// TIA Portal V20 export
ORGANIZATION_BLOCK "T7_Ciclo"   // OB130, LAD, ProgramCycle
TITLE = T7_Ciclo
{ S7_Optimized_Access := 'TRUE' }
AUTHOR : IA
FAMILY : PRUEBA
VERSION : 0.1
// Tanda 3: llama a todas las pruebas
// stored: AutoNumber false, IsIECCheckEnabled false, SetENOAutomatically false
   VAR_INPUT
      Initial_Call : Bool;
      Remanence : Bool;
   END_VAR
BEGIN

REGION Network 1: T7_Base
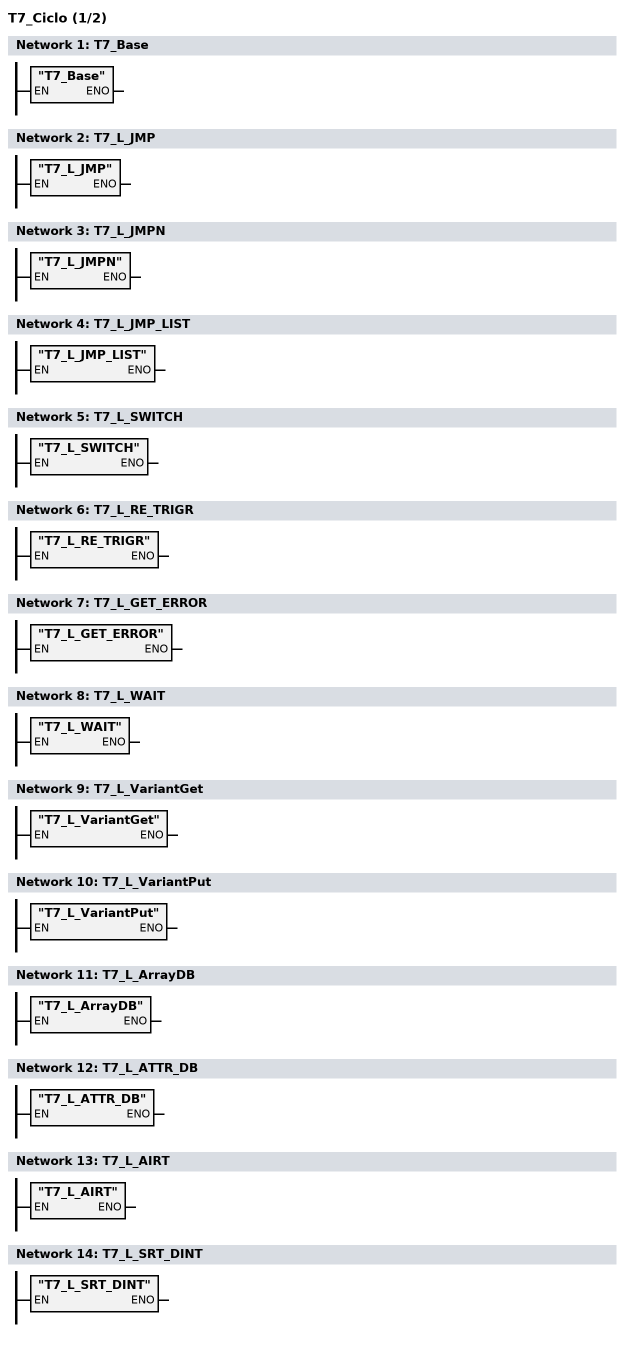
   RUNG wire#powerrail
      "T7_Base"()
   END_RUNG
   // the same network as SCL:
   "T7_Base"();
END_REGION

REGION Network 2: T7_L_JMP
   RUNG wire#powerrail
      "T7_L_JMP"()
   END_RUNG
   // the same network as SCL:
   "T7_L_JMP"();
END_REGION

REGION Network 3: T7_L_JMPN
   RUNG wire#powerrail
      "T7_L_JMPN"()
   END_RUNG
   // the same network as SCL:
   "T7_L_JMPN"();
END_REGION

REGION Network 4: T7_L_JMP_LIST
   RUNG wire#powerrail
      "T7_L_JMP_LIST"()
   END_RUNG
   // the same network as SCL:
   "T7_L_JMP_LIST"();
END_REGION

REGION Network 5: T7_L_SWITCH
   RUNG wire#powerrail
      "T7_L_SWITCH"()
   END_RUNG
   // the same network as SCL:
   "T7_L_SWITCH"();
END_REGION

REGION Network 6: T7_L_RE_TRIGR
   RUNG wire#powerrail
      "T7_L_RE_TRIGR"()
   END_RUNG
   // the same network as SCL:
   "T7_L_RE_TRIGR"();
END_REGION

REGION Network 7: T7_L_GET_ERROR
   RUNG wire#powerrail
      "T7_L_GET_ERROR"()
   END_RUNG
   // the same network as SCL:
   "T7_L_GET_ERROR"();
END_REGION

REGION Network 8: T7_L_WAIT
   RUNG wire#powerrail
      "T7_L_WAIT"()
   END_RUNG
   // the same network as SCL:
   "T7_L_WAIT"();
END_REGION

REGION Network 9: T7_L_VariantGet
   RUNG wire#powerrail
      "T7_L_VariantGet"()
   END_RUNG
   // the same network as SCL:
   "T7_L_VariantGet"();
END_REGION

REGION Network 10: T7_L_VariantPut
   RUNG wire#powerrail
      "T7_L_VariantPut"()
   END_RUNG
   // the same network as SCL:
   "T7_L_VariantPut"();
END_REGION

REGION Network 11: T7_L_ArrayDB
   RUNG wire#powerrail
      "T7_L_ArrayDB"()
   END_RUNG
   // the same network as SCL:
   "T7_L_ArrayDB"();
END_REGION

REGION Network 12: T7_L_ATTR_DB
   RUNG wire#powerrail
      "T7_L_ATTR_DB"()
   END_RUNG
   // the same network as SCL:
   "T7_L_ATTR_DB"();
END_REGION

REGION Network 13: T7_L_AIRT
   RUNG wire#powerrail
      "T7_L_AIRT"()
   END_RUNG
   // the same network as SCL:
   "T7_L_AIRT"();
END_REGION

REGION Network 14: T7_L_SRT_DINT
   RUNG wire#powerrail
      "T7_L_SRT_DINT"()
   END_RUNG
   // the same network as SCL:
   "T7_L_SRT_DINT"();
END_REGION

REGION Network 15: T7_L_QRY_CINT
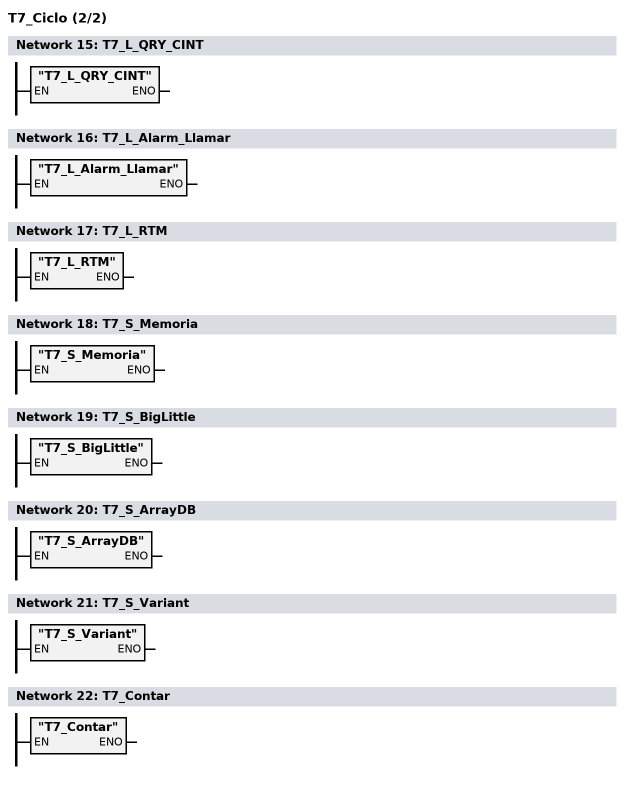
   RUNG wire#powerrail
      "T7_L_QRY_CINT"()
   END_RUNG
   // the same network as SCL:
   "T7_L_QRY_CINT"();
END_REGION

REGION Network 16: T7_L_Alarm_Llamar
   RUNG wire#powerrail
      "T7_L_Alarm_Llamar"()
   END_RUNG
   // the same network as SCL:
   "T7_L_Alarm_Llamar"();
END_REGION

REGION Network 17: T7_L_RTM
   RUNG wire#powerrail
      "T7_L_RTM"()
   END_RUNG
   // the same network as SCL:
   "T7_L_RTM"();
END_REGION

REGION Network 18: T7_S_Memoria
   RUNG wire#powerrail
      "T7_S_Memoria"()
   END_RUNG
   // the same network as SCL:
   "T7_S_Memoria"();
END_REGION

REGION Network 19: T7_S_BigLittle
   RUNG wire#powerrail
      "T7_S_BigLittle"()
   END_RUNG
   // the same network as SCL:
   "T7_S_BigLittle"();
END_REGION

REGION Network 20: T7_S_ArrayDB
   RUNG wire#powerrail
      "T7_S_ArrayDB"()
   END_RUNG
   // the same network as SCL:
   "T7_S_ArrayDB"();
END_REGION

REGION Network 21: T7_S_Variant
   RUNG wire#powerrail
      "T7_S_Variant"()
   END_RUNG
   // the same network as SCL:
   "T7_S_Variant"();
END_REGION

REGION Network 22: T7_Contar
   RUNG wire#powerrail
      "T7_Contar"()
   END_RUNG
   // the same network as SCL:
   "T7_Contar"();
END_REGION
END_ORGANIZATION_BLOCK
